(* IEC 61131-3 sources: iolistgen/tools/tests/fixtures/sample/src/POUs/PRG_Main, 2 files *)

(* ---- PRG_Main.decl.st ---- *)
(*
    Назначение: главная программа — двигатель, выдача выходов, счётчик пусков
    Автор: kr0nsch
    Версия: 1.0.0
    Документ: docs/ARCHITECTURE.md
*)
PROGRAM PRG_Main
VAR
    fbMotor : FB_Motor;
    fbRunEdge : R_TRIG;
    itfDevice : I_Device;
    xInit : BOOL;
END_VAR

(* ---- PRG_Main.impl.st ---- *)
IF NOT xInit THEN
    itfDevice := fbMotor;
    xInit := TRUE;
END_IF

fbMotor(
    stCmd := GVL_Io.stMotorCmd,
    xFeedback := GVL_Io.xMotorFeedback,
    xRun => GVL_Io.xMotorRun);

IF itfDevice <> 0 AND GVL_Io.stMotorCmd.eMode <> itfDevice.Mode THEN
    itfDevice.Mode := GVL_Io.stMotorCmd.eMode;
END_IF

// Счётчик пусков — по фронту события, а не счёт циклов
fbRunEdge(CLK := fbMotor.Running);
IF fbRunEdge.Q THEN
    udiMotorStarts := udiMotorStarts + 1;
END_IF
GVL_Io.stMotorSts := fbMotor.stSts;
